// TIA Portal V20 export
Screen "Pop-up_Mig Weld"  395x500
  ScreenItem "Robot Name" at 2,2 size 393x48  Type=HmiIOField
  ScreenItem "Background" at -1,49 size 395x450  Type=HmiRectangle
  ScreenItem "Cancel Mode" at 315,4 size 76x42  Type=HmiButton
  ScreenItem "矩形_4" at 29,69 size 324x354  Type=HmiRectangle
  ScreenItem "Text Filed E- Stop_17" at 41,345 size 148x21  Type=HmiTextBox
  ScreenItem "Text Field In Auto On_9" at 41,105 size 148x21  Type=HmiTextBox
  ScreenItem "Text Field Home Position_17" at 41,129 size 148x21  Type=HmiTextBox
  ScreenItem "Text field Robot Status_5" at 31,70 size 324x30  Type=HmiTextBox
  ScreenItem "Text Field Manual_17" at 41,273 size 148x21  Type=HmiTextBox
  ScreenItem "Text Field System Ready_9" at 41,153 size 148x21  Type=HmiTextBox
  ScreenItem "Text Field Motor On_9" at 41,177 size 148x21  Type=HmiTextBox
  ScreenItem "Text Field In Cycle_9" at 41,201 size 148x21  Type=HmiTextBox
  ScreenItem "Text Field Cycle On_17" at 41,225 size 148x21  Type=HmiTextBox
  ScreenItem "Text Field On Path_17" at 41,249 size 148x21  Type=HmiTextBox
  ScreenItem "Text Field Tryout Mode_17" at 41,297 size 148x21  Type=HmiTextBox
  ScreenItem "Text Field Stop_17" at 41,321 size 148x21  Type=HmiTextBox
  ScreenItem "Text Filed Error_9" at 41,369 size 148x21  Type=HmiTextBox
  ScreenItem "Text Filed Process Fault_9" at 41,393 size 148x21  Type=HmiTextBox
  ScreenItem "Text Field Home Position_18" at 196,105 size 148x21  Type=HmiTextBox
  ScreenItem "Text Filed E- Stop_18" at 196,249 size 148x21  Type=HmiTextBox
  ScreenItem "Text Field Manual_18" at 196,177 size 148x21  Type=HmiTextBox
  ScreenItem "Text Field Cycle On_18" at 196,129 size 148x21  Type=HmiTextBox
  ScreenItem "Text Field On Path_18" at 196,153 size 148x21  Type=HmiTextBox
  ScreenItem "Text Field Tryout Mode_18" at 196,201 size 148x21  Type=HmiTextBox
  ScreenItem "Text Field Stop_18" at 196,225 size 148x21  Type=HmiTextBox
  ScreenItem "Text Field In Auto On_10" at 196,273 size 148x21  Type=HmiTextBox
  ScreenItem "Text Field Home Position_19" at 196,297 size 148x21  Type=HmiTextBox
  ScreenItem "Text Field System Ready_10" at 196,321 size 148x21  Type=HmiTextBox
  ScreenItem "Text Field Motor On_10" at 196,345 size 148x21  Type=HmiTextBox
  ScreenItem "Text Field Motor On_1" at 196,392 size 148x21  Type=HmiTextBox
  ScreenItem "Text Filed Error_1" at 196,368 size 148x21  Type=HmiTextBox
